(* IEC 61131-3 sources: WenQuest/textbook/plc/ch15/code, 6 files *)

(* ---- p15_3_1.st ---- *)
(* 程序 15.3.1  压装工位的状态机：只有自动循环（方式与异常处理在 15.4、15.5 节加上） *)
TYPE E_Press : (IDLE, CLAMPING, PRESSING, RETURNING, UNCLAMPING); END_TYPE

PROGRAM Main
  VAR
    state : E_Press := IDLE;   (* 当前状态 *)
    tTwoHand : TON;            (* 双手按钮须在 0.5 s 内先后按下 *)
    force : REAL;              (* 压装力，kN *)
    peak : REAL;               (* 本件的最大压装力，kN *)
    resOk, resNok : BOOL;      (* 本件结果：合格 / 不合格 *)
  END_VAR

  force := INT_TO_REAL(AI_Force) * 10.0 / 27648.0;
  tTwoHand(IN := S_Hand1 OR S_Hand2, PT := T#500ms);

  (* 1. 转移：每个状态只看“离开这个状态”的条件 *)
  CASE state OF
    IDLE:
      IF B_Part AND B_PressUp AND B_Unclamped AND S_LC AND S_EStop
         AND S_Hand1 AND S_Hand2 AND NOT tTwoHand.Q THEN
        resOk := FALSE; resNok := FALSE; peak := 0.0;
        state := CLAMPING;
      END_IF;
    CLAMPING:
      IF B_Clamped THEN state := PRESSING; END_IF;
    PRESSING:
      peak := MAX(peak, force);
      IF B_PressDown THEN                          (* 压到底：按最大压装力判定 *)
        resOk := peak >= 4.0 AND peak <= 7.0; resNok := NOT resOk;
        state := RETURNING;
      ELSIF force > 8.0 THEN                       (* 过载：中止，判不合格 *)
        resNok := TRUE; state := RETURNING;
      ELSIF NOT (S_Hand1 AND S_Hand2 AND S_LC) THEN (* 松手或挡光：中止 *)
        resNok := TRUE; state := RETURNING;
      END_IF;
    RETURNING:
      IF B_PressUp THEN state := UNCLAMPING; END_IF;
    UNCLAMPING:
      IF B_Unclamped THEN state := IDLE; END_IF;
  END_CASE;

  (* 2. 输出：只由状态决定，每个输出只写一次 *)
  Y_Clamp     := state = CLAMPING OR state = PRESSING OR state = RETURNING;
  Y_PressDown := state = PRESSING AND S_Hand1 AND S_Hand2 AND S_LC;
  Y_PressUp   := state = RETURNING AND NOT Y_PressDown;   (* 软件联锁：两个线圈不同时得电 *)
  H_OK  := resOk;
  H_NOK := resNok;
  H_Ready := state = IDLE AND B_PressUp AND B_Unclamped;
END_PROGRAM

(* ---- p15_4_1.st ---- *)
(* 程序 15.4.1  压装工位：自动、手动（点动）、单步与回原点 *)
TYPE E_Press : (INIT, HOMING, IDLE, CLAMPING, PRESSING, RETURNING, UNCLAMPING); END_TYPE

PROGRAM Main
  VAR
    state : E_Press := INIT;   (* 上电时位置未知 *)
    auto : BOOL;               (* 自动方式（方式开关在“自动”） *)
    go : BOOL;                 (* 本次扫描允许转移：自动方式下总允许，手动方式下按一次“单步”允许一次 *)
    jog : BOOL;                (* 允许点动：手动方式且停在原点 *)
    rStep, rReset : R_TRIG;
    tTwoHand : TON;
    force, peak : REAL;
    resOk, resNok : BOOL;
  END_VAR

  force := INT_TO_REAL(AI_Force) * 10.0 / 27648.0;
  tTwoHand(IN := S_Hand1 OR S_Hand2, PT := T#500ms);
  rStep(CLK := S_Step);
  rReset(CLK := S_Reset);
  auto := S_Auto;
  go := auto OR rStep.Q;

  CASE state OF
    INIT:                                 (* 等操作员按复位，绝不自己动 *)
      IF rReset.Q AND S_EStop THEN state := HOMING; END_IF;
    HOMING:                               (* 回原点：压头回上位、夹具松开 *)
      IF B_PressUp AND B_Unclamped THEN state := IDLE; END_IF;
    IDLE:
      IF rReset.Q THEN
        state := HOMING;
      ELSIF B_Part AND B_PressUp AND B_Unclamped AND S_LC AND S_EStop
            AND ((auto AND S_Hand1 AND S_Hand2 AND NOT tTwoHand.Q) OR (NOT auto AND rStep.Q)) THEN
        resOk := FALSE; resNok := FALSE; peak := 0.0;
        state := CLAMPING;
      ELSIF NOT auto AND (S_JogClamp OR S_JogDown OR S_JogUp) THEN
        state := INIT;                    (* 点动过：位置不再确定，再启动前要回原点 *)
      END_IF;
    CLAMPING:
      IF go AND B_Clamped THEN state := PRESSING; END_IF;
    PRESSING:
      peak := MAX(peak, force);
      IF force > 8.0 THEN                           (* 过载：任何方式下都立即回程 *)
        resNok := TRUE; state := RETURNING;
      ELSIF go AND B_PressDown THEN
        resOk := peak >= 4.0 AND peak <= 7.0; resNok := NOT resOk;
        state := RETURNING;
      ELSIF auto AND NOT (S_Hand1 AND S_Hand2 AND S_LC) THEN
        resNok := TRUE; state := RETURNING;         (* 自动方式松手或挡光：中止；单步时只是停住 *)
      END_IF;
    RETURNING:
      IF go AND B_PressUp THEN state := UNCLAMPING; END_IF;
    UNCLAMPING:
      IF go AND B_Unclamped THEN state := IDLE; END_IF;
  END_CASE;

  jog := NOT auto AND (state = IDLE OR state = INIT);

  Y_Clamp     := state = CLAMPING OR state = PRESSING OR state = RETURNING OR (jog AND S_JogClamp);
  Y_PressDown := ((state = PRESSING AND S_Hand1 AND S_Hand2) OR (jog AND S_JogDown AND B_Clamped)) AND S_LC AND S_EStop;
  Y_PressUp   := (state = RETURNING OR (state = HOMING AND NOT B_PressUp) OR (jog AND S_JogUp))
                 AND S_EStop AND NOT Y_PressDown;
  H_OK  := resOk;
  H_NOK := resNok;
  H_Ready := state = IDLE;
END_PROGRAM

(* ---- p15_5_1.st ---- *)
(* 程序 15.5.1  压装工位：加上异常处理——动作超时、传感器冲突、急停与恢复 *)
TYPE E_Press : (INIT, HOMING, IDLE, CLAMPING, PRESSING, RETURNING, UNCLAMPING, FAULT, ESTOP); END_TYPE

PROGRAM Main
  VAR
    state : E_Press := INIT;
    prev : E_Press := INIT;    (* 上一次扫描的状态：状态一变，计时重新开始 *)
    tState : TON;              (* 本状态已经停留的时间 *)
    maxTime : TIME;            (* 本状态允许停留的最长时间 *)
    faultCode : INT;               (* 故障代码：0 无；1 夹紧超时；2 压装超时；3 回程超时；4 松开超时；5 回原点超时；9 传感器冲突 *)
    clampHold : BOOL;          (* 进入故障或急停时夹具是否夹着：保持原样 *)
    auto, go, jog : BOOL;
    rStep, rReset : R_TRIG;
    tTwoHand : TON;
    force, peak : REAL;
    resOk, resNok : BOOL;
  END_VAR

  force := INT_TO_REAL(AI_Force) * 10.0 / 27648.0;
  tTwoHand(IN := S_Hand1 OR S_Hand2, PT := T#500ms);
  rStep(CLK := S_Step);
  rReset(CLK := S_Reset);
  auto := S_Auto;
  go := auto OR rStep.Q;

  (* 1. 急停与传感器冲突：任何状态下都优先 *)
  IF NOT S_EStop AND state <> ESTOP THEN
    clampHold := Y_Clamp; state := ESTOP;
  ELSIF ((B_Clamped AND B_Unclamped) OR (B_PressUp AND B_PressDown)) AND state <> FAULT AND state <> ESTOP THEN
    clampHold := Y_Clamp; faultCode := 9; state := FAULT;
  END_IF;

  (* 2. 状态时限：自动方式和回原点时才计时（单步时等的是人） *)
  CASE state OF
    CLAMPING, UNCLAMPING: maxTime := T#1s;
    PRESSING: maxTime := T#4s;
    RETURNING: maxTime := T#5s;
    HOMING: maxTime := T#5s;
  ELSE
    maxTime := T#1h;
  END_CASE;
  tState(IN := state = prev AND (auto OR state = HOMING), PT := maxTime);
  prev := state;

  (* 3. 转移 *)
  CASE state OF
    INIT:
      IF rReset.Q THEN state := HOMING; END_IF;
    HOMING:
      IF B_PressUp AND B_Unclamped THEN state := IDLE;
      ELSIF tState.Q THEN clampHold := FALSE; faultCode := 5; state := FAULT; END_IF;
    IDLE:
      IF rReset.Q THEN
        state := HOMING;
      ELSIF B_Part AND B_PressUp AND B_Unclamped AND S_LC
            AND ((auto AND S_Hand1 AND S_Hand2 AND NOT tTwoHand.Q) OR (NOT auto AND rStep.Q)) THEN
        resOk := FALSE; resNok := FALSE; peak := 0.0;
        state := CLAMPING;
      ELSIF NOT auto AND (S_JogClamp OR S_JogDown OR S_JogUp) THEN
        state := INIT;                    (* 点动过：位置不再确定，再启动前要回原点 *)
      END_IF;
    CLAMPING:
      IF go AND B_Clamped THEN state := PRESSING;
      ELSIF tState.Q THEN clampHold := TRUE; faultCode := 1; state := FAULT; END_IF;
    PRESSING:
      peak := MAX(peak, force);
      IF force > 8.0 THEN
        resNok := TRUE; state := RETURNING;
      ELSIF go AND B_PressDown THEN
        resOk := peak >= 4.0 AND peak <= 7.0; resNok := NOT resOk;
        state := RETURNING;
      ELSIF auto AND NOT (S_Hand1 AND S_Hand2 AND S_LC) THEN
        resNok := TRUE; state := RETURNING;
      ELSIF tState.Q THEN clampHold := TRUE; faultCode := 2; state := FAULT; END_IF;
    RETURNING:
      IF go AND B_PressUp THEN state := UNCLAMPING;
      ELSIF tState.Q THEN clampHold := TRUE; faultCode := 3; state := FAULT; END_IF;
    UNCLAMPING:
      IF go AND B_Unclamped THEN state := IDLE;
      ELSIF tState.Q THEN clampHold := FALSE; faultCode := 4; state := FAULT; END_IF;
    FAULT:                                (* 停在原地，等人看清原因、按复位 *)
      IF rReset.Q AND S_EStop AND NOT ((B_Clamped AND B_Unclamped) OR (B_PressUp AND B_PressDown)) THEN
        faultCode := 0; state := HOMING;
      END_IF;
    ESTOP:                                (* 急停松开后也不自己动，按复位才回原点 *)
      IF S_EStop AND rReset.Q THEN state := HOMING; END_IF;
  END_CASE;

  (* 4. 输出 *)
  jog := NOT auto AND (state = IDLE OR state = INIT OR state = FAULT);   (* 故障时允许点动，联锁照样有效 *)
  Y_Clamp     := state = CLAMPING OR state = PRESSING OR state = RETURNING OR (jog AND S_JogClamp)
                 OR ((state = FAULT OR state = ESTOP) AND clampHold);
  Y_PressDown := ((state = PRESSING AND S_Hand1 AND S_Hand2) OR (jog AND S_JogDown AND B_Clamped)) AND S_LC AND S_EStop;
  Y_PressUp   := (state = RETURNING OR (state = HOMING AND NOT B_PressUp) OR (jog AND S_JogUp))
                 AND S_EStop AND NOT Y_PressDown;
  H_OK    := resOk;
  H_NOK   := resNok;
  H_Ready := state = IDLE;
  H_Fault := state = FAULT OR state = ESTOP;
END_PROGRAM

(* ---- p15_6_1.st ---- *)
(* 程序 15.6.1  三层电梯：用 CASE 写的状态机（呼梯登记、关门、运行、平层、开门） *)
TYPE E_Lift : (DOOR_OPEN, CLOSING, MOVING); END_TYPE

PROGRAM Main
  VAR
    state : E_Lift := DOOR_OPEN;
    call : ARRAY[1..3] OF BOOL;   (* 已登记的呼梯 *)
    floor : INT := 1;             (* 最近经过的楼层 *)
    target : INT;                 (* 要去的楼层，0 表示没有 *)
    tClose : TON;                 (* 关门时限：门被挡住就重新开门 *)
    atTarget : BOOL;
  END_VAR

  (* 登记呼梯；记住最近经过的楼层 *)
  IF S_C1 THEN call[1] := TRUE; END_IF;
  IF S_C2 THEN call[2] := TRUE; END_IF;
  IF S_C3 THEN call[3] := TRUE; END_IF;
  IF B_F1 THEN floor := 1; ELSIF B_F2 THEN floor := 2; ELSIF B_F3 THEN floor := 3; END_IF;
  atTarget := (target = 1 AND B_F1) OR (target = 2 AND B_F2) OR (target = 3 AND B_F3);

  CASE state OF
    DOOR_OPEN:                                   (* 停在某层、门开着 *)
      IF B_F1 OR B_F2 OR B_F3 THEN call[floor] := FALSE; END_IF;   (* 本层的呼梯随到随消 *)
      target := 0;
      IF call[1] THEN target := 1; ELSIF call[2] THEN target := 2; ELSIF call[3] THEN target := 3; END_IF;
      IF target <> 0 AND B_DoorOpen THEN state := CLOSING; END_IF;
    CLOSING:
      tClose(IN := TRUE, PT := T#4s);
      IF B_DoorClosed THEN tClose(IN := FALSE); state := MOVING;
      ELSIF tClose.Q THEN tClose(IN := FALSE); state := DOOR_OPEN; END_IF;
    MOVING:
      IF atTarget THEN call[target] := FALSE; state := DOOR_OPEN; END_IF;
  END_CASE;

  K_Up    := state = MOVING AND target > floor AND NOT atTarget AND S_TopLim AND B_DoorClosed;
  K_Down  := state = MOVING AND target < floor AND NOT atTarget AND S_LowLim AND B_DoorClosed AND NOT K_Up;
  Y_DoorOpen  := state = DOOR_OPEN AND NOT B_DoorOpen;
  Y_DoorClose := state = CLOSING AND NOT B_DoorClosed;
  H_C1 := call[1]; H_C2 := call[2]; H_C3 := call[3];
END_PROGRAM

(* ---- p15_6_2.st ---- *)
(* 程序 15.6.2  三层电梯的顺序功能图写法：同一套 I/O、同样的测试 *)
PROGRAM Main
  VAR
    call : ARRAY[1..3] OF BOOL;
    floor : INT := 1;
    target : INT;
    atTarget : BOOL;
  END_VAR

  IF S_C1 THEN call[1] := TRUE; END_IF;
  IF S_C2 THEN call[2] := TRUE; END_IF;
  IF S_C3 THEN call[3] := TRUE; END_IF;
  IF B_F1 THEN floor := 1; ELSIF B_F2 THEN floor := 2; ELSIF B_F3 THEN floor := 3; END_IF;
  atTarget := (target = 1 AND B_F1) OR (target = 2 AND B_F2) OR (target = 3 AND B_F3);
  H_C1 := call[1]; H_C2 := call[2]; H_C3 := call[3];

  INITIAL_STEP Open: OpenDoor(N); Choose(N); END_STEP
  STEP Closing: Y_DoorClose(N); END_STEP
  STEP Moving: Drive(N); END_STEP
  STEP Arrive: Arrived(P); END_STEP

  ACTION OpenDoor:
    Y_DoorOpen := NOT B_DoorOpen;
  END_ACTION
  ACTION Choose:
    IF B_F1 OR B_F2 OR B_F3 THEN call[floor] := FALSE; END_IF;
    target := 0;
    IF call[1] THEN target := 1; ELSIF call[2] THEN target := 2; ELSIF call[3] THEN target := 3; END_IF;
  END_ACTION
  ACTION Drive:
    K_Up   := target > floor AND NOT atTarget AND S_TopLim AND B_DoorClosed;
    K_Down := target < floor AND NOT atTarget AND S_LowLim AND B_DoorClosed AND NOT K_Up;
  END_ACTION
  ACTION Arrived:
    K_Up := FALSE; K_Down := FALSE; call[target] := FALSE;
  END_ACTION

  TRANSITION FROM Open TO Closing := target <> 0 AND B_DoorOpen; END_TRANSITION
  TRANSITION FROM Closing TO Moving := B_DoorClosed; END_TRANSITION
  TRANSITION FROM Closing TO Open := Closing.T >= T#4s; END_TRANSITION       (* 门被挡住：重新开门 *)
  TRANSITION FROM Moving TO Arrive := atTarget; END_TRANSITION
  TRANSITION FROM Arrive TO Open := TRUE; END_TRANSITION
END_PROGRAM

(* ---- p15_7_1.st ---- *)
(* 程序 15.7.1  错误的做法：把状态变量设成保持型（RETAIN）。其余与程序 15.5.1 完全相同 *)
TYPE E_Press : (INIT, HOMING, IDLE, CLAMPING, PRESSING, RETURNING, UNCLAMPING, FAULT, ESTOP); END_TYPE

PROGRAM Main
  VAR RETAIN                   (* ← 断电后保持 *)
    state : E_Press := INIT;
    prev : E_Press := INIT;
  END_VAR
  VAR
    tState : TON;              (* 本状态已经停留的时间 *)
    maxTime : TIME;            (* 本状态允许停留的最长时间 *)
    faultCode : INT;               (* 故障代码：0 无；1 夹紧超时；2 压装超时；3 回程超时；4 松开超时；5 回原点超时；9 传感器冲突 *)
    clampHold : BOOL;          (* 进入故障或急停时夹具是否夹着：保持原样 *)
    auto, go, jog : BOOL;
    rStep, rReset : R_TRIG;
    tTwoHand : TON;
    force, peak : REAL;
    resOk, resNok : BOOL;
  END_VAR

  force := INT_TO_REAL(AI_Force) * 10.0 / 27648.0;
  tTwoHand(IN := S_Hand1 OR S_Hand2, PT := T#500ms);
  rStep(CLK := S_Step);
  rReset(CLK := S_Reset);
  auto := S_Auto;
  go := auto OR rStep.Q;

  (* 1. 急停与传感器冲突：任何状态下都优先 *)
  IF NOT S_EStop AND state <> ESTOP THEN
    clampHold := Y_Clamp; state := ESTOP;
  ELSIF ((B_Clamped AND B_Unclamped) OR (B_PressUp AND B_PressDown)) AND state <> FAULT AND state <> ESTOP THEN
    clampHold := Y_Clamp; faultCode := 9; state := FAULT;
  END_IF;

  (* 2. 状态时限：自动方式和回原点时才计时（单步时等的是人） *)
  CASE state OF
    CLAMPING, UNCLAMPING: maxTime := T#1s;
    PRESSING: maxTime := T#4s;
    RETURNING: maxTime := T#5s;
    HOMING: maxTime := T#5s;
  ELSE
    maxTime := T#1h;
  END_CASE;
  tState(IN := state = prev AND (auto OR state = HOMING), PT := maxTime);
  prev := state;

  (* 3. 转移 *)
  CASE state OF
    INIT:
      IF rReset.Q THEN state := HOMING; END_IF;
    HOMING:
      IF B_PressUp AND B_Unclamped THEN state := IDLE;
      ELSIF tState.Q THEN clampHold := FALSE; faultCode := 5; state := FAULT; END_IF;
    IDLE:
      IF rReset.Q THEN
        state := HOMING;
      ELSIF B_Part AND B_PressUp AND B_Unclamped AND S_LC
            AND ((auto AND S_Hand1 AND S_Hand2 AND NOT tTwoHand.Q) OR (NOT auto AND rStep.Q)) THEN
        resOk := FALSE; resNok := FALSE; peak := 0.0;
        state := CLAMPING;
      ELSIF NOT auto AND (S_JogClamp OR S_JogDown OR S_JogUp) THEN
        state := INIT;                    (* 点动过：位置不再确定，再启动前要回原点 *)
      END_IF;
    CLAMPING:
      IF go AND B_Clamped THEN state := PRESSING;
      ELSIF tState.Q THEN clampHold := TRUE; faultCode := 1; state := FAULT; END_IF;
    PRESSING:
      peak := MAX(peak, force);
      IF force > 8.0 THEN
        resNok := TRUE; state := RETURNING;
      ELSIF go AND B_PressDown THEN
        resOk := peak >= 4.0 AND peak <= 7.0; resNok := NOT resOk;
        state := RETURNING;
      ELSIF auto AND NOT (S_Hand1 AND S_Hand2 AND S_LC) THEN
        resNok := TRUE; state := RETURNING;
      ELSIF tState.Q THEN clampHold := TRUE; faultCode := 2; state := FAULT; END_IF;
    RETURNING:
      IF go AND B_PressUp THEN state := UNCLAMPING;
      ELSIF tState.Q THEN clampHold := TRUE; faultCode := 3; state := FAULT; END_IF;
    UNCLAMPING:
      IF go AND B_Unclamped THEN state := IDLE;
      ELSIF tState.Q THEN clampHold := FALSE; faultCode := 4; state := FAULT; END_IF;
    FAULT:                                (* 停在原地，等人看清原因、按复位 *)
      IF rReset.Q AND S_EStop AND NOT ((B_Clamped AND B_Unclamped) OR (B_PressUp AND B_PressDown)) THEN
        faultCode := 0; state := HOMING;
      END_IF;
    ESTOP:                                (* 急停松开后也不自己动，按复位才回原点 *)
      IF S_EStop AND rReset.Q THEN state := HOMING; END_IF;
  END_CASE;

  (* 4. 输出 *)
  jog := NOT auto AND (state = IDLE OR state = INIT OR state = FAULT);   (* 故障时允许点动，联锁照样有效 *)
  Y_Clamp     := state = CLAMPING OR state = PRESSING OR state = RETURNING OR (jog AND S_JogClamp)
                 OR ((state = FAULT OR state = ESTOP) AND clampHold);
  Y_PressDown := ((state = PRESSING AND S_Hand1 AND S_Hand2) OR (jog AND S_JogDown AND B_Clamped)) AND S_LC AND S_EStop;
  Y_PressUp   := (state = RETURNING OR (state = HOMING AND NOT B_PressUp) OR (jog AND S_JogUp))
                 AND S_EStop AND NOT Y_PressDown;
  H_OK    := resOk;
  H_NOK   := resNok;
  H_Ready := state = IDLE;
  H_Fault := state = FAULT OR state = ESTOP;
END_PROGRAM
